(* IEC 61131-3 sources: rusty/tests/lit/cfc/blocks/action_call, 2 files *)

(* ---- main.st ---- *)
FUNCTION main : DINT
    action_call();
    action_call();
    // CHECK: count = 6
    printf('count = %d$N', action_call.result);
END_FUNCTION

(* ---- counter.st ---- *)
FUNCTION_BLOCK counter
VAR_INPUT
    step : DINT;
END_VAR
VAR_OUTPUT
    count : DINT;
END_VAR
END_FUNCTION_BLOCK

ACTIONS
    ACTION bump
        count := count + step;
    END_ACTION
END_ACTIONS
